// TIA Portal V20 export
VAR_GLOBAL   // PLC tag table "STEP7 classic symbols"
END_VAR
